Fanuc KAREL source: KA00216.KL

PROGRAM KA00216
%NOLOCKGROUP
VAR
  SRC: ARRAY[4] OF XYZWPR
  DST: ARRAY[4] OF JOINTPOS
BEGIN
  DST = SRC
END KA00216
